Staubli VAL3: getArmTypeList.pgx

public program getArmTypeList(string& x_sItem[], string& x_sItem2[])
// //获取所有4轴6轴机器人型号列表
// //x_sItem  4轴手臂型号列表
// //x_sItem2 6轴手臂型号列表
  local trsf l_tTrsf
  local string l_sItem[6]
  local string l_sEvent
  local string l_sItem2[7]
  local string l_sKey[2]
  local num i
  local num j
begin
  //获取所有4轴6轴机器人型号列表
  //x_sItem  4轴手臂型号列表
  //x_sItem2 6轴手臂型号列表
  //获取列表
  resize(x_sItem,1,size(forcedata:tArm4Force))
  resize(x_sItem2,1,size(forcedata:tArm6Force))
  l_sKey=first(forcedata:tArm4Force)
  l_sKey[1]=first(forcedata:tArm6Force)
  i=0
  j=0
  while l_sKey!=""
    x_sItem[i]=l_sKey
    l_sKey=next(forcedata:tArm4Force[l_sKey])
    i=i+1
  endWhile
  while l_sKey[1]!=""
    x_sItem2[j]=l_sKey[1]
    l_sKey[1]=next(forcedata:tArm6Force[l_sKey[1]])
    j=j+1
  endWhile
  if l_sKey=="" and i==0
    x_sItem[i]=""
  endIf
  if l_sKey[1]=="" and j==0
    x_sItem2[j]=""
  endIf
end
